(* IEC 61131-3 sources: plcassist-cli/packages/volt-lsp-iec/test-corpus/pro2193/Device/Plc Logic/Application/09 Misc/Library Manager/(unresolved)/cmpusermgr implementation, 51 files *)

(* ---- USERMGRCHANGEMYPASSWORD.fun ---- *)
FUNCTION USERMGRCHANGEMYPASSWORD : RTS_IEC_RESULT
VAR_INPUT
	HUSER : RTS_IEC_HANDLE;
	PSZUSER : REFERENCE TO STRING;
	PSZOLDPASSWORD : REFERENCE TO STRING;
	PSZNEWPASSWORD : REFERENCE TO STRING;
END_VAR
END_FUNCTION

(* ---- USERMGRGETSESSIONUSER.fun ---- *)
FUNCTION USERMGRGETSESSIONUSER : RTS_IEC_HANDLE
VAR_INPUT
	SESSIONID : UDINT;
	PRESULT : POINTER TO RTS_IEC_RESULT;
END_VAR
END_FUNCTION

(* ---- USERMGRGETUSERACCESSRIGHTS.fun ---- *)
FUNCTION USERMGRGETUSERACCESSRIGHTS : RTS_IEC_RESULT
VAR_INPUT
	PSZOBJECT : REFERENCE TO STRING;
	HUSER : RTS_IEC_HANDLE;
	PULRIGHTS : POINTER TO DWORD;
	PULDENIEDRIGHTS : POINTER TO DWORD;
END_VAR
END_FUNCTION

(* ---- USERMGRGROUPADD.fun ---- *)
FUNCTION USERMGRGROUPADD : RTS_IEC_RESULT
VAR_INPUT
	HUSER : RTS_IEC_HANDLE;
END_VAR
VAR_IN_OUT
	PSZGROUPNAME : STRING;
END_VAR
END_FUNCTION

(* ---- USERMGRGROUPADDUSER.fun ---- *)
FUNCTION USERMGRGROUPADDUSER : RTS_IEC_RESULT
VAR_INPUT
	HUSER : RTS_IEC_HANDLE;
END_VAR
VAR_IN_OUT
	PSZGROUPNAME : STRING;
	PSZUSERNAME : STRING;
END_VAR
END_FUNCTION

(* ---- USERMGRGROUPGETFIRST.fun ---- *)
FUNCTION USERMGRGROUPGETFIRST : RTS_IEC_HANDLE
VAR_INPUT
	HUSER : RTS_IEC_HANDLE;
END_VAR
VAR_OUTPUT
	RESULT : RTS_IEC_RESULT;
END_VAR
END_FUNCTION

(* ---- USERMGRGROUPGETFIRSTUSER.fun ---- *)
FUNCTION USERMGRGROUPGETFIRSTUSER : RTS_IEC_RESULT
VAR_INPUT
	HUSER : RTS_IEC_HANDLE;
	HGROUP : RTS_IEC_HANDLE;
END_VAR
VAR_IN_OUT
	PHITERATOR : RTS_IEC_HANDLE;
	PSZUSERNAME : STRING(59);
END_VAR
END_FUNCTION

(* ---- USERMGRGROUPGETFIRSTUSERINTERNAL.fun ---- *)
FUNCTION USERMGRGROUPGETFIRSTUSERINTERNAL : RTS_IEC_RESULT
VAR_INPUT
	HUSER : RTS_IEC_HANDLE;
	HGROUP : RTS_IEC_HANDLE;
	IMAXLEN : UDINT;
END_VAR
VAR_IN_OUT
	PHITERATOR : RTS_IEC_HANDLE;
	PSZUSERNAME : STRING;
END_VAR
END_FUNCTION

(* ---- USERMGRGROUPGETHANDLE.fun ---- *)
FUNCTION USERMGRGROUPGETHANDLE : RTS_IEC_HANDLE
VAR_INPUT
	HUSER : RTS_IEC_HANDLE;
END_VAR
VAR_OUTPUT
	RESULT : RTS_IEC_RESULT;
END_VAR
VAR_IN_OUT
	PSZGROUPNAME : STRING;
END_VAR
END_FUNCTION

(* ---- USERMGRGROUPGETNAME.fun ---- *)
FUNCTION USERMGRGROUPGETNAME : RTS_IEC_RESULT
VAR_INPUT
	HUSER : RTS_IEC_HANDLE;
	HGROUP : RTS_IEC_HANDLE;
END_VAR
VAR_IN_OUT
	PSZGROUP : STRING(59);
END_VAR
END_FUNCTION

(* ---- USERMGRGROUPGETNAMEINTERNAL.fun ---- *)
FUNCTION USERMGRGROUPGETNAMEINTERNAL : RTS_IEC_RESULT
VAR_INPUT
	HUSER : RTS_IEC_HANDLE;
	HGROUP : RTS_IEC_HANDLE;
	IMAXLEN : UDINT;
END_VAR
VAR_IN_OUT
	PSZGROUP : STRING;
END_VAR
END_FUNCTION

(* ---- USERMGRGROUPGETNEXT.fun ---- *)
FUNCTION USERMGRGROUPGETNEXT : RTS_IEC_HANDLE
VAR_INPUT
	HUSER : RTS_IEC_HANDLE;
	HPREVGROUP : RTS_IEC_HANDLE;
END_VAR
VAR_OUTPUT
	RESULT : RTS_IEC_RESULT;
END_VAR
END_FUNCTION

(* ---- USERMGRGROUPGETNEXTUSER.fun ---- *)
FUNCTION USERMGRGROUPGETNEXTUSER : RTS_IEC_RESULT
VAR_INPUT
	HUSER : RTS_IEC_HANDLE;
	HGROUP : RTS_IEC_HANDLE;
END_VAR
VAR_IN_OUT
	PHITERATOR : RTS_IEC_HANDLE;
	PSZUSERNAME : STRING(59);
END_VAR
END_FUNCTION

(* ---- USERMGRGROUPGETNEXTUSERINTERNAL.fun ---- *)
FUNCTION USERMGRGROUPGETNEXTUSERINTERNAL : RTS_IEC_RESULT
VAR_INPUT
	HUSER : RTS_IEC_HANDLE;
	HGROUP : RTS_IEC_HANDLE;
	IMAXLEN : UDINT;
END_VAR
VAR_IN_OUT
	PHITERATOR : RTS_IEC_HANDLE;
	PSZUSERNAME : STRING;
END_VAR
END_FUNCTION

(* ---- USERMGRGROUPREMOVE.fun ---- *)
FUNCTION USERMGRGROUPREMOVE : RTS_IEC_RESULT
VAR_INPUT
	HUSER : RTS_IEC_HANDLE;
END_VAR
VAR_IN_OUT
	PSZGROUPNAME : STRING;
END_VAR
END_FUNCTION

(* ---- USERMGRGROUPREMOVEUSER.fun ---- *)
FUNCTION USERMGRGROUPREMOVEUSER : RTS_IEC_RESULT
VAR_INPUT
	HUSER : RTS_IEC_HANDLE;
END_VAR
VAR_IN_OUT
	PSZGROUP : STRING;
	PSZUSER : STRING;
END_VAR
END_FUNCTION

(* ---- USERMGRHASUSERACCESSRIGHTS.fun ---- *)
FUNCTION USERMGRHASUSERACCESSRIGHTS : RTS_IEC_RESULT
VAR_INPUT
	PSZOBJECT : REFERENCE TO STRING;
	HUSER : RTS_IEC_HANDLE;
	ULREQUESTEDRIGHTS : DWORD;
END_VAR
END_FUNCTION

(* ---- USERMGRISACTIVE.fun ---- *)
FUNCTION USERMGRISACTIVE : BOOL
END_FUNCTION

(* ---- USERMGRLOGIN.fun ---- *)
FUNCTION USERMGRLOGIN : RTS_IEC_HANDLE
VAR_INPUT
	PSZUSER : REFERENCE TO STRING;
	PSZPASSWORD : REFERENCE TO STRING;
	PRESULT : POINTER TO RTS_IEC_RESULT;
END_VAR
END_FUNCTION

(* ---- USERMGRLOGOUT.fun ---- *)
FUNCTION USERMGRLOGOUT : RTS_IEC_RESULT
VAR_INPUT
	HUSER : RTS_IEC_HANDLE;
END_VAR
END_FUNCTION

(* ---- USERMGROBJECTADD.fun ---- *)
FUNCTION USERMGROBJECTADD : RTS_IEC_HANDLE
VAR_INPUT
	PSZOBJECT : REFERENCE TO STRING;
	PRESULT : POINTER TO RTS_IEC_RESULT;
END_VAR
END_FUNCTION

(* ---- USERMGROBJECTADDGROUP.fun ---- *)
FUNCTION USERMGROBJECTADDGROUP : RTS_IEC_RESULT
VAR_INPUT
	HUSER : RTS_IEC_HANDLE;
	HOBJECT : RTS_IEC_HANDLE;
	HGROUP : RTS_IEC_HANDLE;
END_VAR
END_FUNCTION

(* ---- USERMGROBJECTCLEARRIGHTS.fun ---- *)
FUNCTION USERMGROBJECTCLEARRIGHTS : RTS_IEC_RESULT
VAR_INPUT
	HUSER : RTS_IEC_HANDLE;
	HOBJECT : RTS_IEC_HANDLE;
END_VAR
END_FUNCTION

(* ---- USERMGROBJECTGETFIRSTCHILD.fun ---- *)
FUNCTION USERMGROBJECTGETFIRSTCHILD : RTS_IEC_HANDLE
VAR_INPUT
	HFATHEROBJECT : RTS_IEC_HANDLE;
END_VAR
VAR_OUTPUT
	RESULT : RTS_IEC_RESULT;
END_VAR
END_FUNCTION

(* ---- USERMGROBJECTGETFIRSTGROUP.fun ---- *)
FUNCTION USERMGROBJECTGETFIRSTGROUP : RTS_IEC_HANDLE
VAR_INPUT
	HUSER : RTS_IEC_HANDLE;
	HOBJECT : RTS_IEC_HANDLE;
END_VAR
VAR_OUTPUT
	RESULT : RTS_IEC_RESULT;
END_VAR
END_FUNCTION

(* ---- USERMGROBJECTGETGROUPRIGHTS.fun ---- *)
FUNCTION USERMGROBJECTGETGROUPRIGHTS : RTS_IEC_RESULT
VAR_INPUT
	HUSER : RTS_IEC_HANDLE;
	HOBJECT : RTS_IEC_HANDLE;
	HGROUP : RTS_IEC_HANDLE;
END_VAR
VAR_OUTPUT
	ULRIGHTS : DWORD;
	ULDENIEDRIGHTS : DWORD;
END_VAR
END_FUNCTION

(* ---- USERMGROBJECTGETHANDLE.fun ---- *)
FUNCTION USERMGROBJECTGETHANDLE : RTS_IEC_HANDLE
VAR_OUTPUT
	RESULT : RTS_IEC_RESULT;
END_VAR
VAR_IN_OUT
	PSZOBJECTNAME : STRING;
END_VAR
END_FUNCTION

(* ---- USERMGROBJECTGETNAME.fun ---- *)
FUNCTION USERMGROBJECTGETNAME : RTS_IEC_RESULT
VAR_INPUT
	HOBJECT : RTS_IEC_HANDLE;
	PSZOBJECT : POINTER TO STRING;
	PIMAXLEN : POINTER TO UDINT;
END_VAR
END_FUNCTION

(* ---- USERMGROBJECTGETNEXTCHILD.fun ---- *)
FUNCTION USERMGROBJECTGETNEXTCHILD : RTS_IEC_HANDLE
VAR_INPUT
	HFATHEROBJECT : RTS_IEC_HANDLE;
	HPREVCHILD : RTS_IEC_HANDLE;
END_VAR
VAR_OUTPUT
	RESULT : RTS_IEC_RESULT;
END_VAR
END_FUNCTION

(* ---- USERMGROBJECTGETNEXTGROUP.fun ---- *)
FUNCTION USERMGROBJECTGETNEXTGROUP : RTS_IEC_HANDLE
VAR_INPUT
	HUSER : RTS_IEC_HANDLE;
	HOBJECT : RTS_IEC_HANDLE;
	HPREVGROUP : RTS_IEC_HANDLE;
END_VAR
VAR_OUTPUT
	RESULT : RTS_IEC_RESULT;
END_VAR
END_FUNCTION

(* ---- USERMGROBJECTREMOVE.fun ---- *)
FUNCTION USERMGROBJECTREMOVE : RTS_IEC_RESULT
VAR_INPUT
	HOBJECT : RTS_IEC_HANDLE;
END_VAR
END_FUNCTION

(* ---- USERMGROBJECTREMOVEGROUP.fun ---- *)
FUNCTION USERMGROBJECTREMOVEGROUP : RTS_IEC_RESULT
VAR_INPUT
	HUSER : RTS_IEC_HANDLE;
	HOBJECT : RTS_IEC_HANDLE;
	HGROUP : RTS_IEC_HANDLE;
END_VAR
END_FUNCTION

(* ---- USERMGROBJECTSETGROUPDENIEDRIGHTS.fun ---- *)
FUNCTION USERMGROBJECTSETGROUPDENIEDRIGHTS : RTS_IEC_RESULT
VAR_INPUT
	HUSER : RTS_IEC_HANDLE;
	HOBJECT : RTS_IEC_HANDLE;
	HGROUP : RTS_IEC_HANDLE;
	ULDENIEDRIGHTS : DWORD;
END_VAR
END_FUNCTION

(* ---- USERMGROBJECTSETGROUPRIGHTS.fun ---- *)
FUNCTION USERMGROBJECTSETGROUPRIGHTS : RTS_IEC_RESULT
VAR_INPUT
	HUSER : RTS_IEC_HANDLE;
	HOBJECT : RTS_IEC_HANDLE;
	HGROUP : RTS_IEC_HANDLE;
	ULRIGHTS : DWORD;
END_VAR
END_FUNCTION

(* ---- USERMGROBJECTSETUSEDRIGHTS.fun ---- *)
FUNCTION USERMGROBJECTSETUSEDRIGHTS : RTS_IEC_RESULT
VAR_INPUT
	HOBJECT : RTS_IEC_HANDLE;
	ULUSEDRIGHTS : DWORD;
END_VAR
END_FUNCTION

(* ---- USERMGRRELOGIN.fun ---- *)
FUNCTION USERMGRRELOGIN : RTS_IEC_RESULT
VAR_INPUT
	HUSER : RTS_IEC_HANDLE;
	PSZUSER : REFERENCE TO STRING;
	PSZPASSWORD : REFERENCE TO STRING;
END_VAR
END_FUNCTION

(* ---- USERMGRUSERADD.fun ---- *)
FUNCTION USERMGRUSERADD : RTS_IEC_RESULT
VAR_INPUT
	HUSER : RTS_IEC_HANDLE;
END_VAR
VAR_IN_OUT
	PSZUSER : STRING;
	PCREDENTIALS : UserMgrCredentials;
END_VAR
END_FUNCTION

(* ---- USERMGRUSERADDINFOTOUSER.fun ---- *)
FUNCTION USERMGRUSERADDINFOTOUSER : RTS_IEC_RESULT
VAR_INPUT
	HUSER : RTS_IEC_HANDLE;
	KEY : __XWORD;
	VALUE : UserMgrCacheValue;
END_VAR
END_FUNCTION

(* ---- USERMGRUSERGETFIRST.fun ---- *)
FUNCTION USERMGRUSERGETFIRST : RTS_IEC_RESULT
VAR_INPUT
	HUSER : RTS_IEC_HANDLE;
END_VAR
VAR_OUTPUT
	USERPROPERTY : DWORD;
END_VAR
VAR_IN_OUT
	PHITERATOR : RTS_IEC_HANDLE;
	PSZUSERNAME : STRING(59);
END_VAR
END_FUNCTION

(* ---- USERMGRUSERGETFIRSTINTERNAL.fun ---- *)
FUNCTION USERMGRUSERGETFIRSTINTERNAL : RTS_IEC_RESULT
VAR_INPUT
	HUSER : RTS_IEC_HANDLE;
	IMAXLEN : UDINT;
END_VAR
VAR_OUTPUT
	USERPROPERTY : DWORD;
END_VAR
VAR_IN_OUT
	PHITERATOR : RTS_IEC_HANDLE;
	PSZUSERNAME : STRING;
END_VAR
END_FUNCTION

(* ---- USERMGRUSERGETINFOOFUSER.fun ---- *)
FUNCTION USERMGRUSERGETINFOOFUSER : DWORD
VAR_INPUT
	HUSER : RTS_IEC_HANDLE;
	KEY : __XWORD;
END_VAR
VAR_OUTPUT
	VALUE : UserMgrCacheValue;
END_VAR
END_FUNCTION

(* ---- USERMGRUSERGETNAME.fun ---- *)
FUNCTION USERMGRUSERGETNAME : RTS_IEC_RESULT
VAR_INPUT
	HUSER : RTS_IEC_HANDLE;
END_VAR
VAR_IN_OUT
	PSZUSERNAME : STRING(59);
END_VAR
END_FUNCTION

(* ---- USERMGRUSERGETNAMEINTERNAL.fun ---- *)
FUNCTION USERMGRUSERGETNAMEINTERNAL : RTS_IEC_RESULT
VAR_INPUT
	HUSER : RTS_IEC_HANDLE;
	IMAXLEN : UDINT;
END_VAR
VAR_IN_OUT
	PSZUSERNAME : STRING;
END_VAR
END_FUNCTION

(* ---- USERMGRUSERGETNEXT.fun ---- *)
FUNCTION USERMGRUSERGETNEXT : RTS_IEC_RESULT
VAR_INPUT
	HUSER : RTS_IEC_HANDLE;
END_VAR
VAR_OUTPUT
	USERPROPERTY : DWORD;
END_VAR
VAR_IN_OUT
	PHITERATOR : RTS_IEC_HANDLE;
	PSZUSERNAME : STRING(59);
END_VAR
END_FUNCTION

(* ---- USERMGRUSERGETNEXTINTERNAL.fun ---- *)
FUNCTION USERMGRUSERGETNEXTINTERNAL : RTS_IEC_RESULT
VAR_INPUT
	HUSER : RTS_IEC_HANDLE;
	IMAXLEN : UDINT;
END_VAR
VAR_OUTPUT
	USERPROPERTY : DWORD;
END_VAR
VAR_IN_OUT
	PHITERATOR : RTS_IEC_HANDLE;
	PSZUSERNAME : STRING;
END_VAR
END_FUNCTION

(* ---- USERMGRUSERGETPROPERTY.fun ---- *)
FUNCTION USERMGRUSERGETPROPERTY : DWORD
VAR_INPUT
	HUSER : RTS_IEC_HANDLE;
END_VAR
VAR_OUTPUT
	RESULT : RTS_IEC_RESULT;
END_VAR
VAR_IN_OUT
	PSZUSER : STRING;
END_VAR
END_FUNCTION

(* ---- USERMGRUSERREMOVE.fun ---- *)
FUNCTION USERMGRUSERREMOVE : RTS_IEC_RESULT
VAR_INPUT
	HUSER : RTS_IEC_HANDLE;
END_VAR
VAR_IN_OUT
	PSZUSER : STRING;
END_VAR
END_FUNCTION

(* ---- USERMGRUSERREMOVEINFOFROMALLUSERS.fun ---- *)
FUNCTION USERMGRUSERREMOVEINFOFROMALLUSERS : DWORD
VAR_INPUT
	KEY : __XWORD;
END_VAR
END_FUNCTION

(* ---- USERMGRUSERREMOVEINFOFROMUSER.fun ---- *)
FUNCTION USERMGRUSERREMOVEINFOFROMUSER : DWORD
VAR_INPUT
	HUSER : RTS_IEC_HANDLE;
	KEY : __XWORD;
END_VAR
END_FUNCTION

(* ---- USERMGRUSERSETCREDENTIALS.fun ---- *)
FUNCTION USERMGRUSERSETCREDENTIALS : RTS_IEC_RESULT
VAR_INPUT
	HUSER : RTS_IEC_HANDLE;
END_VAR
VAR_IN_OUT
	PSZUSER : STRING;
	PCREDENTIALS : UserMgrCredentials;
END_VAR
END_FUNCTION

(* ---- USERMGRUSERSETPROPERTY.fun ---- *)
FUNCTION USERMGRUSERSETPROPERTY : RTS_IEC_RESULT
VAR_INPUT
	HUSER : RTS_IEC_HANDLE;
	USERPROPERTY : DWORD;
END_VAR
VAR_IN_OUT
	PSZUSER : STRING;
END_VAR
END_FUNCTION
